FUNCTION_BLOCK SortingSequence1 (* Composite Function Block Type *)
  (* Standard: 61499-2 *)
  (* Version 0.0, 7/2/2026, template *)
  PACKAGE Main;
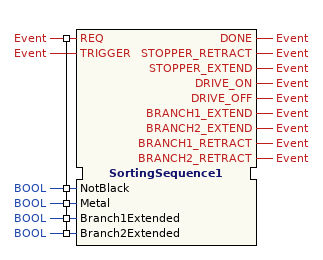
  EVENT_INPUT
    REQ WITH NotBlack, Metal, Branch1Extended, Branch2Extended; (* Normal Execution Request *)
    TRIGGER;
  END_EVENT
  EVENT_OUTPUT
    DONE; (* Initialization Confirm *)
    STOPPER_RETRACT; (* Execution Confirmation *)
    STOPPER_EXTEND;
    DRIVE_ON;
    DRIVE_OFF;
    BRANCH1_EXTEND;
    BRANCH2_EXTEND;
    BRANCH1_RETRACT;
    BRANCH2_RETRACT;
  END_EVENT
  VAR_INPUT
    NotBlack : BOOL; (* Input event qualifier *)
    Metal : BOOL;
    Branch1Extended : BOOL;
    Branch2Extended : BOOL;
  END_VAR
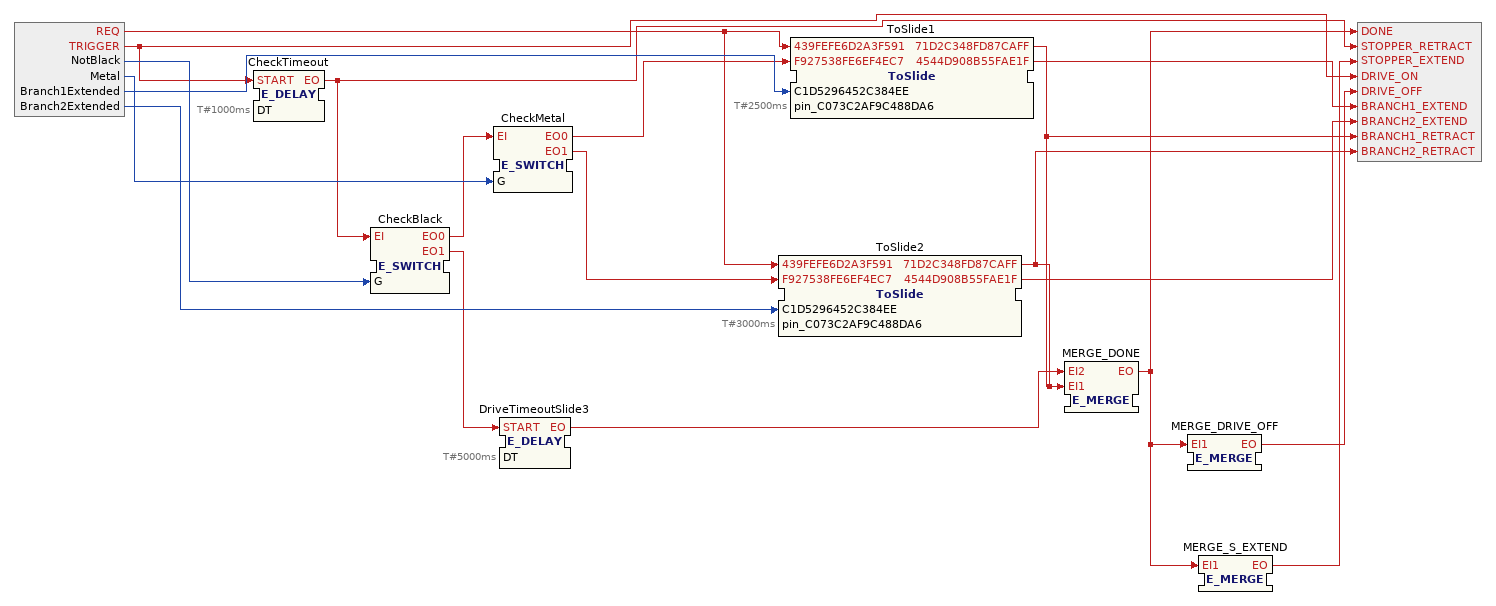
  FBS
    CheckTimeout : E_DELAY(DT := T#1000ms);
    DriveTimeoutSlide3 : E_DELAY(DT := T#5000ms);
    CheckBlack : E_SWITCH;
    CheckMetal : E_SWITCH;
    ToSlide1 : ToSlide(pin_C073C2AF9C488DA6 := T#2500ms);
    ToSlide2 : ToSlide(pin_C073C2AF9C488DA6 := T#3000ms);
    MERGE_DONE : E_MERGE;
    MERGE_DRIVE_OFF : E_MERGE;
    MERGE_S_EXTEND : E_MERGE;
  END_FBS
  EVENT_CONNECTIONS
    TRIGGER TO CheckTimeout.START;
    TRIGGER TO DRIVE_ON;
    REQ TO ToSlide1.439FEFE6D2A3F591;
    REQ TO ToSlide2.439FEFE6D2A3F591;
    CheckTimeout.EO TO CheckBlack.EI;
    CheckTimeout.EO TO STOPPER_RETRACT;
    CheckBlack.EO0 TO CheckMetal.EI;
    CheckBlack.EO1 TO DriveTimeoutSlide3.START;
    CheckMetal.EO0 TO ToSlide1.F927538FE6EF4EC7;
    CheckMetal.EO1 TO ToSlide2.F927538FE6EF4EC7;
    DriveTimeoutSlide3.EO TO MERGE_DONE.EI2;
    MERGE_DONE.EO TO MERGE_S_EXTEND.EI1;
    MERGE_DONE.EO TO MERGE_DRIVE_OFF.EI1;
    MERGE_DRIVE_OFF.EO TO DRIVE_OFF;
    MERGE_S_EXTEND.EO TO STOPPER_EXTEND;
    MERGE_DONE.EO TO DONE;
    ToSlide1.71D2C348FD87CAFF TO MERGE_DONE.EI1;
    ToSlide1.71D2C348FD87CAFF TO BRANCH1_RETRACT;
    ToSlide2.71D2C348FD87CAFF TO MERGE_DONE.EI1;
    ToSlide2.71D2C348FD87CAFF TO BRANCH2_RETRACT;
    ToSlide1.4544D908B55FAE1F TO BRANCH1_EXTEND;
    ToSlide2.4544D908B55FAE1F TO BRANCH2_EXTEND;
  END_CONNECTIONS
  DATA_CONNECTIONS
    NotBlack TO CheckBlack.G;
    Metal TO CheckMetal.G;
    Branch2Extended TO ToSlide2.C1D5296452C384EE;
    Branch1Extended TO ToSlide1.C1D5296452C384EE;
  END_CONNECTIONS
END_FUNCTION_BLOCK
